Staubli VAL3: safeZoneCheck.pgx

public program safeZoneCheck()
  local bool l_bResult
  local bool l_bErr
  local num l_i
begin
  for l_i = 0 to size(safeTemp:zZoneItem)-1
    if safeTemp:zZoneItem[l_i].bActive
      call computeZone(l_i,l_bResult)
      call io:setDigOutput(O_safeZone[l_i],l_bResult,l_bErr)
    endIf
  endFor
end
